(* IEC 61131-3 sources: Caravan/Archiv/12-04-19/Stations/MachineControl/MachineControl/Network/Licht_Net, 1 file *)

(* ---- ONE_Licht_Net_Table.st ---- *)
#define OBJECTS_CONFIG

FUNCTION GLOBAL TAB ONE_Licht_Net
-1$UINT, 0$UINT,
0$UINT, 0$UINT,

1$UDINT,
TO_UDINT(2856325874), "NightLight_Class", 0$UINT, 0$UINT, 1$UINT,

_NO_ATTR, TO_UDINT(3502587029), "NIGHTLIGHT_CLASS1",

//Internal connections
0$UDINT,
0$UDINT,
0$UDINT,
0$UDINT,

//Initialization values
0$UDINT,
1$UDINT,
TO_UDINT(0), "OC_To_Timer_Class", TO_UDINT(0),//|Licht_Net.NightLight_Class1.OC_To_Timer_Class;

//Symbolic initialization values
0$UDINT,
0$UDINT,

//Initialization of string values
0$UDINT,
0$UDINT,

//Configuration of tasks (RealTime, Cyclic, Background)
0$UDINT,
0$UDINT,

0$UDINT,
1$UDINT,
TO_UDINT(0), (-2147483598)$UDINT, 4194303$DINT, 	//NIGHTLIGHT_CLASS1

0$UDINT,
0$UDINT,

//External connections
0$UDINT,
2$UDINT,
TO_UDINT(0), "OC_To_Timer_Class", C_DIR, TO_UDINT(1302809437), "Timer_Class1","ClassSvr",
TO_UDINT(0), "cNightlightSwitch", C_DIR, TO_UDINT(542619847), "SR0201","Led350",

//Magic internal connections
0$UDINT,
0$UDINT,

//Configuration of timeslots of tasks (RealTime, Cyclic)
#ifdef __LSLLDR_TIMESLOTS__
0$UDINT,
0$UDINT,

0$UDINT,
0$UDINT,

#endif //__LSLLDR_TIMESLOTS__

//MultiMaster connections
#ifdef __LSLLDR_MULTIMASTER__
0$UDINT,
0$UDINT,
#endif //__LSLLDR_MULTIMASTER__

//Configuration for task ID (RealTime, CyclicTime)
#ifdef __LSLLDR_TASKID__
"\\\\TASKS2  "
0$UDINT,
0$UDINT,

0$UDINT,
1$UDINT,
(0)$UDINT, 	//NIGHTLIGHT_CLASS1

0$UDINT,
0$UDINT,

#endif //__LSLLDR_TASKID__

END_FUNCTION
